VISUALIZATION Screen2  // 2x2
END_VISUALIZATION

(* stored: Version 1.1.0.1, ProductVersion 3.1.4024.15
   Visu Screen2: Id {2f7f4d1c-2d56-4174-a889-f22cd0bf7f28} *)
